Fanuc KAREL source: KO00069.KL

PROGRAM KO00069
%NOLOCKGROUP
%ENVIRONMENT MIR
VAR
  P1: XYZWPREXT
  P2: XYZWPR
  F: BOOLEAN
  OUT: POSITION
BEGIN
  F = TRUE
  OUT = MIRROR(P1, P2, F)
END KO00069
